// TIA Portal V21 export
Screen "T02_RectApp"  1024x768, Number=22
  ScreenLayer 
    Rectangle "P_CellRect" at 0,0 size 100x30
      AppearanceAnimation   AnimationMode=Range, Tag=CellSt0_00
        AppearanceAnimationRange 
        AppearanceAnimationRange   Range=1
        AppearanceAnimationRange   Range=2
        AppearanceAnimationRange   Range=3
        AppearanceAnimationRange   Range=4
        AppearanceAnimationRange   Range=5
        AppearanceAnimationRange   Range=6
        AppearanceAnimationRange   Range=7
